// TIA Portal V21 export
// export: Created 2026-10-23T20:43:30.4071431Z, ExportSetting WithDefaults, DisplayName Totally Integrated Automation Portal, DisplayVersion V21 Update 1, DisplayName SINAMICS Startdrive Advanced, DisplayVersion V21 HF2, DisplayName SINAMICS Startdrive G110M, G120, G120C, G120D, G120P, G115D, DisplayVersion V21 HF2, DisplayName SINAMICS Startdrive G130, G150, S120, S150, G200, G220, S200, S210, S220, Innomotics MVD, DisplayVersion V21 HF2, DisplayName STEP 7 Professional, DisplayVersion V21 Update 1, DisplayName STEP 7 Safety, DisplayVersion V21, DisplayName Tech WebApplication, DisplayVersion V21, DisplayName WinCC Basic/Comfort/Advanced, DisplayVersion V21 Update 1, DisplayName WinCC Unified, DisplayVersion V21 Update 1
FUNCTION_BLOCK "FB_AnaStatusIgnored"   // FB18, SCL
TITLE = Analyzer: status never evaluated
{ S7_Optimized_Access := 'TRUE' }
VERSION : 0.1
// Rule C26n: RET_VAL of RD_LOC_T is stored but never evaluated
// stored: AutoNumber true, IsIECCheckEnabled false, IsRetainMemResEnabled false, MemoryReserve 100, SetENOAutomatically false, UDAEnableTagReadback false
   VAR
      Now : DTL;   // Local time
   END_VAR
   VAR_TEMP
      RetVal : Int;   // Status of RD_LOC_T
   END_VAR
BEGIN

       #RetVal := RD_LOC_T(OUT => #Now);
END_FUNCTION_BLOCK
